(* IEC 61131-3 sources: codesys-api/examples/plc_architecture/st, 45 files *)

(* ---- E_BusFormat.st ---- *)
// How an entry's raw value sits in a block's reply: one bit, or one or two 16-bit registers.
{attribute 'qualified_only'}
{attribute 'strict'}
TYPE E_BusFormat :
(
	SINGLE_BIT := 0,
	INT16 := 1,
	UINT16 := 2,
	INT32 := 3,
	UINT32 := 4,
	FLOAT32 := 5
) USINT;
END_TYPE

(* ---- E_BusFunction.st ---- *)
// Modbus read function of a poll block. Writes (FC06) come from GVL_Bus.Writes.
{attribute 'qualified_only'}
{attribute 'strict'}
TYPE E_BusFunction :
(
	READ_COILS := 1,
	READ_DISCRETE_INPUTS := 2,
	READ_HOLDING_REGISTERS := 3,
	READ_INPUT_REGISTERS := 4
) USINT;
END_TYPE

(* ---- E_CommandResult.st ---- *)
// Outcome of a remote command, sent back to the sender in the acknowledgement. A retry of an id the PLC has
// already answered gets the original result again; it is never applied twice.
{attribute 'qualified_only'}
{attribute 'strict'}
TYPE E_CommandResult :
(
	PENDING := 0,           // parsed, not yet checked
	ACCEPTED := 1,
	MALFORMED := 2,         // not "<id>,<tag>=<number>,<sent_ms>", or a field too long
	UNKNOWN_TAG := 3,
	NOT_WRITABLE := 4,
	OUT_OF_RANGE := 5,      // outside the tag's range, not 0/1 for a BOOL, not whole for an INT, NaN
	TOO_OLD := 6,           // older than allowed, dated in the future, or waited too long in the queue
	OUT_OF_ORDER := 7,      // older than the last command applied to the same tag
	INTERLOCKED := 8,       // a start while not permitted, or sent before the permit came back
	CLOCK_NOT_SYNCED := 9   // the PLC's wall clock isn't plausible, so freshness can't be checked
) USINT;
END_TYPE

(* ---- E_Quality.st ---- *)
// Quality of a tag's value. Interlocks and publishing look at this, not just at the number.
{attribute 'qualified_only'}
{attribute 'strict'}
TYPE E_Quality :
(
	INIT := 0,          // no value since start-up
	GOOD := 1,
	STALE := 2,         // no fresh value from the source within StaleAfter
	COMM_FAIL := 3,     // the source reports a communication error
	INVALID := 4        // out of range, or not computable (e.g. division by zero)
) USINT;
END_TYPE

(* ---- E_TagKind.st ---- *)
{attribute 'qualified_only'}
{attribute 'strict'}
TYPE E_TagKind :
(
	BOOL_TAG := 0,
	INT_TAG := 1,
	REAL_TAG := 2
) USINT;
END_TYPE

(* ---- ST_BusBlock.st ---- *)
// One read request, repeated every PeriodMs: a run of registers or bits of one device. The generator merges a
// device's nearby channels into as few blocks as possible (at most 125 registers or 2,000 bits each).
TYPE ST_BusBlock :
STRUCT
	Line : INT;                         // index in GVL_Bus.Lines
	UnitId : UINT;
	ReadFunction : E_BusFunction;
	Start : UINT;                       // zero-based register or bit address (CODESYS numbering)
	Count : UINT;
	PeriodMs : UDINT := 1000;
	FirstEntry : INT;                   // GVL_Bus.Entries[FirstEntry .. FirstEntry + EntryCount - 1]
	EntryCount : INT;
	Source : INT;                       // the device's source in GVL_Tags (health and age)
END_STRUCT
END_TYPE

(* ---- ST_BusEntry.st ---- *)
// Where one tag's raw value sits in its block's reply. Scaling is the tag's own (ST_TagConfig.Scale and
// Offset); the bus only delivers the device's number.
TYPE ST_BusEntry :
STRUCT
	Offset : UINT;                      // registers (or bits) from the block's Start
	Format : E_BusFormat;
	IsWordSwapped : BOOL;               // 32-bit values: low word first
	HasSentinel : BOOL;                 // a raw value the device uses for "no reading"
	Sentinel : DINT;                    // e.g. -999 for an open thermocouple; delivered as NaN, so the tag is INVALID
	TagIndex : INT;
END_STRUCT
END_TYPE

(* ---- ST_BusLine.st ---- *)
// One Modbus connection: a TCP server (a device or an RS485 gateway port) or one of the PLC's serial ports.
// Every device on it shares this one connection; requests on it run one at a time.
TYPE ST_BusLine :
STRUCT
	IsSerial : BOOL;
	Address : ARRAY[0..3] OF BYTE;      // TCP: server IP
	Port : UINT := 502;                 // TCP: server port
	ComPort : INT := 1;                 // serial: 1 to 4
	RtsControl : USINT;                 // serial: 0 disabled, 1 on, 2 handshake, 3 toggle (RS485 direction)
	Baudrate : UDINT := 9600;           // serial: 9600, 19200, 38400, 57600 or 115200
	Parity : USINT;                     // serial: 0 none, 1 odd, 2 even
	ReplyTimeoutMs : UDINT := 500;
END_STRUCT
END_TYPE

(* ---- ST_BusWrite.st ---- *)
// A writable tag sent to a device register (FC06) when its value changes, and again every RefreshMs so a
// device that restarted gets it back. Raw = (Value - tag Offset) / tag Scale, as a signed 16-bit register.
TYPE ST_BusWrite :
STRUCT
	TagIndex : INT;                     // 0 = unused row
	Line : INT;
	UnitId : UINT;
	Register : UINT;
	RefreshMs : UDINT := 10000;
END_STRUCT
END_TYPE

(* ---- ST_Command.st ---- *)
// One remote command, from the MQTT callback to the control task and back as an acknowledgement.
TYPE ST_Command :
STRUCT
	Id : UDINT;                 // sender's command id, echoed in the acknowledgement
	TagIndex : INT;             // resolved when received; 0 = unknown tag
	Value : REAL;
	SentAtMs : ULINT;           // wall-clock ms from the bridge, the one command sender
	ReceivedAtMs : ULINT;
	Result : E_CommandResult;
END_STRUCT
END_TYPE

(* ---- ST_TagConfig.st ---- *)
// Static description of one tag. Generated from the config sheet into GVL_Tags.TagConfig;
// the program never writes it.
TYPE ST_TagConfig :
STRUCT
	Name : STRING(24);          // tag key, exactly as the bridge layout spells it; sized by the generator from the longest name
	Kind : E_TagKind;
	Scale : REAL := 1.0;        // Value := Raw * Scale + Offset
	Offset : REAL;
	MinValue : REAL;            // a value outside [MinValue, MaxValue], or NaN, is INVALID
	MaxValue : REAL;
	DefaultValue : REAL;        // writable tags start here (alarm setpoints from the sheet; requests 0)
	Deadband : REAL;            // report-by-exception: publish when the value moved more than this
	StaleAfter : TIME := T#5S;  // no fresh value from the source for this long -> STALE
	IsWritable : BOOL;          // may a remote command change it (setpoints, start/stop requests)?
	Source : INT;               // communication source in GVL_Tags.SourceIsHealthy; 0 = local I/O
END_STRUCT
END_TYPE

(* ---- ST_TagState.st ---- *)
// Live state of one tag. Written only by PRG_Control, each field by one step.
TYPE ST_TagState :
STRUCT
	Raw : REAL;                 // step 1: as read from the I/O or the bus
	SourceQuality : E_Quality;  // step 1: from the source's health and age
	Value : REAL;               // step 3 (step 2 for writable tags); BOOL tags use 0.0 / 1.0
	Quality : E_Quality;        // step 3: SourceQuality plus range checks (step 2 for writable tags)
	UpdatedAtMs : ULINT;        // step 1 (step 2 for writable tags): last fresh value, monotonic ms
	LastCommandSentAtMs : ULINT; // step 2: sender time of the last command applied, for ordering
END_STRUCT
END_TYPE

(* ---- GVL_Bus.st ---- *)
// Modbus devices and their hand-over to the control task. Tables are generated from the config sheets'
// rs485Config (and Modbus TCP devices); PRG_Bus (bus task) is the only writer of everything below them.
// Example: AIT-1508 is holding register 40002 (item 1) of RTU unit 24 on the PLC's first serial port.
{attribute 'qualified_only'}
VAR_GLOBAL CONSTANT
	LINE_COUNT : INT := 1;
	BLOCK_COUNT : INT := 1;
	ENTRY_COUNT : INT := 1;
	WRITE_COUNT : INT := 1;
	FAIL_LIMIT : UINT := 3;             // consecutive failed requests before a device is COMM_FAIL
	BACKOFF_MS : UDINT := 5000;         // a failed device is polled this rarely, so it can't slow its line
END_VAR
VAR_GLOBAL
	// Generated; never written by the program.
	Lines : ARRAY[1..LINE_COUNT] OF ST_BusLine := [(IsSerial := TRUE, ComPort := 1, Baudrate := 9600)];
	Blocks : ARRAY[1..BLOCK_COUNT] OF ST_BusBlock := [
		(Line := 1, UnitId := 24, ReadFunction := E_BusFunction.READ_HOLDING_REGISTERS, Start := 1, Count := 1,
		 PeriodMs := 500, FirstEntry := 1, EntryCount := 1, Source := 1)];
	Entries : ARRAY[1..ENTRY_COUNT] OF ST_BusEntry := [(Offset := 0, Format := E_BusFormat.UINT16, TagIndex := 1)];
	Writes : ARRAY[1..WRITE_COUNT] OF ST_BusWrite;          // no device setpoints in this example
	IsBusSource : ARRAY[0..GVL_Tags.SOURCE_COUNT] OF BOOL := [FALSE, TRUE, FALSE];

	// Bus task -> control task. For a source with SourceWriting TRUE the control task was started while the
	// bus task was mid-update: it keeps last scan's values for that source. (Both tasks on one core: control
	// never runs while the bus task writes, except by preempting it.)
	Raw : ARRAY[1..GVL_Tags.TAG_COUNT] OF REAL;             // decoded device numbers, before tag scaling
	SourceWriting : ARRAY[0..GVL_Tags.SOURCE_COUNT] OF BOOL;
	SourceHealthy : ARRAY[0..GVL_Tags.SOURCE_COUNT] OF BOOL := [TRUE, TRUE, TRUE];   // until FAIL_LIMIT failures: INIT, not COMM_FAIL
	SourceLastGoodMs : ARRAY[0..GVL_Tags.SOURCE_COUNT] OF ULINT;   // F_NowMs of the last good reply

	// Diagnostics
	SourceFailCount : ARRAY[0..GVL_Tags.SOURCE_COUNT] OF UINT;
	BlockReads : ARRAY[1..BLOCK_COUNT] OF UDINT;
	BlockErrors : ARRAY[1..BLOCK_COUNT] OF UDINT;
	BlockLastError : ARRAY[1..BLOCK_COUNT] OF UDINT;        // ModbusFB.Error
	BlockLastException : ARRAY[1..BLOCK_COUNT] OF UDINT;    // Modbus exception code
	WriteCount : ARRAY[1..WRITE_COUNT] OF UDINT;
	WriteErrors : ARRAY[1..WRITE_COUNT] OF UDINT;
END_VAR

(* ---- GVL_Tags.st ---- *)
// The tag table and the hand-over points between the control task and the comms task.
// Ownership: every variable below has exactly one writer, named in its comment.
// Changing the table (rows, order, sizes) needs a full download: queued commands and the publisher's
// history refer to rows by index, so an online change must not reinterpret them.
{attribute 'qualified_only'}
VAR_GLOBAL CONSTANT
	TAG_COUNT : INT := 4;               // generated from the config sheet
	SOURCE_COUNT : INT := 2;            // Modbus slaves and remote PLCs; 0 = local I/O
	// Indices for hand-written logic, generated with the table so names and indices stay in step
	TAG_AIT_1508 : INT := 1;
	TAG_AIT_1508_HH_SP : INT := 2;
	TAG_P_1502_REQUEST : INT := 3;
	TAG_LSS_E_STOP : INT := 4;
END_VAR
VAR_GLOBAL
	// Generated from the config sheet; never written by the program.
	TagConfig : ARRAY[1..TAG_COUNT] OF ST_TagConfig := [
		(Name := 'AIT-1508', Kind := E_TagKind.REAL_TAG, Scale := 0.01, MinValue := 0.0, MaxValue := 14.0,
		 Deadband := 0.05, StaleAfter := T#3S, Source := 1),
		(Name := 'AIT-1508_HH_SP', Kind := E_TagKind.REAL_TAG, MinValue := 0.0, MaxValue := 14.0,
		 DefaultValue := 12.5, IsWritable := TRUE),
		(Name := 'P-1502', Kind := E_TagKind.BOOL_TAG, MinValue := 0.0, MaxValue := 1.0, IsWritable := TRUE),
		(Name := 'LSS-E-STOP', Kind := E_TagKind.BOOL_TAG, MinValue := 0.0, MaxValue := 1.0, StaleAfter := T#3S, Source := 2)];

	Tags : ARRAY[1..TAG_COUNT] OF ST_TagState;               // writer: PRG_Control
	RawInputs : ARRAY[1..TAG_COUNT] OF REAL;                  // writer: I/O mapping (control task)
	// Source health and the time of each source's last sample. Writer: the source adapters, which run in the
	// control task (Modbus diagnostics are read there). Data from other tasks (e.g. remote PLCs over MQTT)
	// reaches them through a queue, never by writing these from another task. Not in the skeleton.
	SourceIsHealthy : ARRAY[0..SOURCE_COUNT] OF BOOL := [TRUE, FALSE, FALSE];
	SourceUpdatedAtMs : ARRAY[0..SOURCE_COUNT] OF ULINT;      // 0 = no sample since start-up

	// Control -> comms: a consistent copy of Tags, made when the comms task asks for one.
	PublishSnapshot : ARRAY[1..TAG_COUNT] OF ST_TagState;    // writer: PRG_Control
	SnapshotRequest : UDINT;                                  // writer: PRG_Comms (increments to ask)
	SnapshotSequence : UDINT;                                 // writer: PRG_Control (= SnapshotRequest when served)

	// Comms -> control and back. Each queue has one producer task and one consumer task.
	// Both tasks must run on the same core, or the queues need the target's atomics and barriers.
	Commands : FB_CommandQueue;         // Push: FB_CommandReceiver (comms task); Pop: PRG_Control
	Acks : FB_CommandQueue;             // Push: PRG_Control; Pop: PRG_Comms

	// Physical outputs, mapped to I/O.
	P_1502_RUN : BOOL;                  // writer: PRG_Control.WriteOutputs, nothing else
END_VAR

(* ---- F_BusDecode.st ---- *)
FUNCTION F_BusDecode : BOOL
// Turns one block's reply into GVL_Bus.Raw for each of its entries. Call it with the source's SourceWriting
// flag set. A sentinel ("no reading") becomes NaN, so the tag goes INVALID in ComputeValues. Independent of
// the transport: FB_BusLine passes a ModbusFB reply, a native device-tree channel its mapped input image.
VAR_INPUT
	FirstEntry : INT;
	EntryCount : INT;
END_VAR
VAR_IN_OUT
	Words : ARRAY[0..124] OF WORD;      // register reply, first register at index 0
	Bits : ARRAY[0..1999] OF BYTE;      // bit reply, one byte per bit
END_VAR
VAR
	Index : INT;
	Entry : ST_BusEntry;
	RawInt : DINT;
	Raw32 : DWORD;
	Value : REAL;
	pReal : POINTER TO REAL;
	NanBits : DWORD := 16#7FC00000;
END_VAR
// ---- implementation ----
FOR Index := FirstEntry TO FirstEntry + EntryCount - 1 DO
	Entry := GVL_Bus.Entries[Index];
	IF Entry.Format = E_BusFormat.SINGLE_BIT THEN
		RawInt := SEL(Bits[Entry.Offset] <> 0, 0, 1);   // ModbusFB unpacks bit replies: one byte per coil (bench, 2026-10-20)
		Value := DINT_TO_REAL(RawInt);
	ELSIF Entry.Format = E_BusFormat.INT16 THEN
		RawInt := INT_TO_DINT(WORD_TO_INT(Words[Entry.Offset]));
		Value := DINT_TO_REAL(RawInt);
	ELSIF Entry.Format = E_BusFormat.UINT16 THEN
		RawInt := WORD_TO_DINT(Words[Entry.Offset]);
		Value := DINT_TO_REAL(RawInt);
	ELSE
		IF Entry.IsWordSwapped THEN
			Raw32 := SHL(WORD_TO_DWORD(Words[Entry.Offset + 1]), 16) OR WORD_TO_DWORD(Words[Entry.Offset]);
		ELSE
			Raw32 := SHL(WORD_TO_DWORD(Words[Entry.Offset]), 16) OR WORD_TO_DWORD(Words[Entry.Offset + 1]);
		END_IF
		RawInt := DWORD_TO_DINT(Raw32);
		IF Entry.Format = E_BusFormat.FLOAT32 THEN
			pReal := ADR(Raw32);
			Value := pReal^;
		ELSIF Entry.Format = E_BusFormat.UINT32 THEN
			Value := UDINT_TO_REAL(DWORD_TO_UDINT(Raw32));
		ELSE
			Value := DINT_TO_REAL(RawInt);
		END_IF
	END_IF
	IF Entry.HasSentinel AND RawInt = Entry.Sentinel THEN
		pReal := ADR(NanBits);
		Value := pReal^;
	END_IF
	GVL_Bus.Raw[Entry.TagIndex] := Value;
END_FOR
F_BusDecode := TRUE;

(* ---- F_FindTag.st ---- *)
FUNCTION F_FindTag : INT
// Index of the tag with this name, 0 if there is none. A linear search is fine for occasional commands;
// with thousands of tags and frequent commands, generate the table sorted by name and search it binarily.
VAR_INPUT
	Name : STRING(24);
END_VAR
VAR
	Index : INT;
END_VAR
// ---- implementation ----
F_FindTag := 0;
FOR Index := 1 TO GVL_Tags.TAG_COUNT DO
	IF GVL_Tags.TagConfig[Index].Name = Name THEN
		F_FindTag := Index;
		RETURN;
	END_IF
END_FOR

(* ---- F_IsNumberText.st ---- *)
FUNCTION F_IsNumberText : BOOL
// TRUE for a plain decimal number of 1..MaxLength characters: an optional leading '-', digits, at most one
// '.'. With IsDigitsOnly, only unsigned integers (ids, timestamps). MaxLength keeps the value inside the
// target type (9 digits for a UDINT id, 15 for a millisecond timestamp). Run this before STRING_TO_REAL/
// _UDINT/_ULINT, which return 0 for text they can't read.
VAR_INPUT
	Text : STRING(40);
	IsDigitsOnly : BOOL;
	MaxLength : INT;
END_VAR
VAR
	pChar : POINTER TO BYTE;
	Length : INT;
	Index : INT;
	Digits : INT;
	Dots : INT;
END_VAR
// ---- implementation ----
F_IsNumberText := FALSE;
Length := LEN(Text);
IF Length < 1 OR Length > MaxLength THEN
	RETURN;
END_IF
pChar := ADR(Text);
FOR Index := 0 TO Length - 1 DO
	IF pChar[Index] >= 16#30 AND pChar[Index] <= 16#39 THEN
		Digits := Digits + 1;
	ELSIF pChar[Index] = 16#2E AND NOT IsDigitsOnly THEN
		Dots := Dots + 1;
	ELSIF NOT (pChar[Index] = 16#2D AND Index = 0 AND NOT IsDigitsOnly) THEN
		RETURN;                         // any other character, or '-' anywhere but first
	END_IF
END_FOR
F_IsNumberText := Digits > 0 AND Dots <= 1;

(* ---- F_NowMs.st ---- *)
FUNCTION F_NowMs : ULINT
// Monotonic milliseconds since start-up, for ages and timeouts. Not wall-clock time.
VAR
	Microseconds : ULINT;
END_VAR
// ---- implementation ----
SysTimeCore.SysTimeGetUs(pUsTime := Microseconds);
F_NowMs := Microseconds / 1000;

(* ---- F_NowUs.st ---- *)
FUNCTION F_NowUs : ULINT
// Monotonic microseconds since start-up, for time budgets within a scan. Not wall-clock time.
VAR
	Microseconds : ULINT;
END_VAR
// ---- implementation ----
SysTimeCore.SysTimeGetUs(pUsTime := Microseconds);
F_NowUs := Microseconds;

(* ---- F_WallClockMs.st ---- *)
FUNCTION F_WallClockMs : ULINT
// Milliseconds since 1970 from the controller's real-time clock, to compare with senders' timestamps.
// Only meaningful while the clock is synchronized (SNTP).
VAR
	Timestamp : ULINT;
END_VAR
// ---- implementation ----
SysTimeRtc.SysTimeRtcHighResGet(pTimestamp := Timestamp);
F_WallClockMs := Timestamp;

(* ---- FB_BusLine.st ---- *)
{attribute 'no_assign'}
FUNCTION_BLOCK FB_BusLine
// One Modbus connection (GVL_Bus.Lines[LineIndex]) with every block and write on it. Called every bus-task
// cycle. One request is in flight at a time; the next starts in the same call that finishes the last
// (ModbusFB's "daisy chain"), so the line never idles a task cycle between requests.
VAR_INPUT
	LineIndex : INT;
	IsEnabled : BOOL := TRUE;
	Reconnect : BOOL;                   // rising edge: drop the connection and connect with the current settings
END_VAR
VAR_OUTPUT
	IsConnected : BOOL;
	RequestCount : UDINT;
	ErrorCount : UDINT;
	LastRequestUs : UDINT;              // start to reply of the last request
	MaxRequestUs : UDINT;
END_VAR
VAR
	ClientTcp : ModbusFB.ClientTCP;
	ClientRtu : ModbusFB.ClientSerial;
	Client : REFERENCE TO ModbusFB.Client;   // whichever of the two this line uses (set by CallClient)
	ReadCoils : ModbusFB.ClientRequestReadCoils;
	ReadDiscrete : ModbusFB.ClientRequestReadDiscreteInputs;
	ReadHolding : ModbusFB.ClientRequestReadHoldingRegisters;
	ReadInput : ModbusFB.ClientRequestReadInputRegisters;
	WriteRegister : ModbusFB.ClientRequestWriteSingleRegister;
	Words : ARRAY[0..124] OF WORD;      // reply of the active register block
	Bits : ARRAY[0..1999] OF BYTE;      // reply of the active bit block: one byte per bit (ModbusFB unpacks them)
	Block : ST_BusBlock;                // copy of the active block
	ActiveBlock : INT;                  // 0 = no read in flight
	ActiveWrite : INT;                  // 0 = no write in flight
	NextBlock : INT := 1;               // round-robin start
	BlockDueMs : ARRAY[1..GVL_Bus.BLOCK_COUNT] OF ULINT;
	WriteDueMs : ARRAY[1..GVL_Bus.WRITE_COUNT] OF ULINT;
	WriteSentValue : ARRAY[1..GVL_Bus.WRITE_COUNT] OF REAL;
	HasWritten : ARRAY[1..GVL_Bus.WRITE_COUNT] OF BOOL;
	WriteValue : REAL;
	WriteRaw : INT;
	IsDone : BOOL;
	IsError : BOOL;
	ErrorId : UDINT;
	Exception : UDINT;
	NowMs : ULINT;
	StartUs : ULINT;
	ReconnectEdge : R_TRIG;
	HoldUntilMs : ULINT;                // connection held down until then (reconnect, client error)
END_VAR
// ---- implementation ----
NowMs := F_NowMs();
ReconnectEdge(CLK := Reconnect);
IF ReconnectEdge.Q THEN
	HoldUntilMs := NowMs + 500;
END_IF
CallClient();

IF ActiveBlock <> 0 OR ActiveWrite <> 0 THEN
	IF CallRequest(IsExecute := TRUE) THEN
		FinishRequest();
	END_IF
END_IF
IF ActiveBlock = 0 AND ActiveWrite = 0 AND IsConnected THEN
	StartNext();
END_IF

(* ---- FB_CommandQueue.st ---- *)
FUNCTION_BLOCK FB_CommandQueue
// Single-producer / single-consumer ring buffer between two tasks. Push is called from one task
// only, Pop from one other task only; each side writes only its own index, so no lock is needed. Push fills
// the slot before it advances Head, so Pop never sees a half-written item. This relies on both tasks running
// on one core; across cores, the index updates need the runtime's atomic operations and memory barriers.
// Usable capacity is SIZE - 1 (one slot stays empty to tell "full" from "empty").
VAR CONSTANT
	SIZE : UINT := 32;
END_VAR
VAR_OUTPUT
	OverflowCount : UDINT;              // items dropped because the queue was full
END_VAR
VAR
	Items : ARRAY[0..SIZE - 1] OF ST_Command;
	Head : UINT;                        // next free slot; written only by Push
	Tail : UINT;                        // next item to take; written only by Pop
END_VAR
// ---- implementation ----
// Everything happens in the Push and Pop methods.

(* ---- FB_CommandReceiver.st ---- *)
FUNCTION_BLOCK FB_CommandReceiver IMPLEMENTS MQTT.MQTT_SUBSCRIBE_CALLBACK
// MQTT subscription callback: turns every received command into an ST_Command and queues it for the
// control task, instead of keeping only the latest message. Runs in the comms task (inside the MQTT client).
// Message format: <id>,<tag>=<value>,<sent_ms>   e.g. '1042,P-1502=1,1769612037947'
VAR_OUTPUT
	ReceivedCount : UDINT;
	MalformedCount : UDINT;
	DroppedCount : UDINT;               // queue full: no acknowledgement, so the sender retries
END_VAR
VAR
	Line : STRING(255);
END_VAR
// ---- implementation ----
// Everything happens in PublishReceived, called by the MQTT library for each message.

(* ---- FB_BusLine.CallClient.st ---- *)
METHOD CallClient : BOOL
// Runs this line's client (TCP or serial) and returns IsConnected. Settings are read when it connects. A client
// error holds the connection down for a second before the next attempt.
VAR
	Port : SysCom.SYS_COM_PORTS;
	Baudrate : SysCom.SYS_COM_BAUDRATE;
	Parity : SysCom.SYS_COM_PARITY;
	Rts : SysCom.SYS_COM_RTS_CONTROL;
END_VAR
// ---- implementation ----
IF GVL_Bus.Lines[LineIndex].IsSerial THEN
	CASE GVL_Bus.Lines[LineIndex].ComPort OF
		2: Port := SysCom.SYS_COM_PORTS.SYS_COMPORT2;
		3: Port := SysCom.SYS_COM_PORTS.SYS_COMPORT3;
		4: Port := SysCom.SYS_COM_PORTS.SYS_COMPORT4;
	ELSE
		Port := SysCom.SYS_COM_PORTS.SYS_COMPORT1;
	END_CASE
	CASE GVL_Bus.Lines[LineIndex].RtsControl OF
		1: Rts := SysCom.SYS_COM_RTS_CONTROL.SYS_RTS_CONTROL_ENABLE;
		2: Rts := SysCom.SYS_COM_RTS_CONTROL.SYS_RTS_CONTROL_HANDSHAKE;
		3: Rts := SysCom.SYS_COM_RTS_CONTROL.SYS_RTS_CONTROL_TOGGLE;
	ELSE
		Rts := SysCom.SYS_COM_RTS_CONTROL.SYS_RTS_CONTROL_DISABLE;
	END_CASE
	CASE GVL_Bus.Lines[LineIndex].Baudrate OF
		19200: Baudrate := SysCom.SYS_COM_BAUDRATE.SYS_BR_19200;
		38400: Baudrate := SysCom.SYS_COM_BAUDRATE.SYS_BR_38400;
		57600: Baudrate := SysCom.SYS_COM_BAUDRATE.SYS_BR_57600;
		115200: Baudrate := SysCom.SYS_COM_BAUDRATE.SYS_BR_115200;
	ELSE
		Baudrate := SysCom.SYS_COM_BAUDRATE.SYS_BR_9600;
	END_CASE
	CASE GVL_Bus.Lines[LineIndex].Parity OF
		1: Parity := SysCom.SYS_COM_PARITY.SYS_ODDPARITY;
		2: Parity := SysCom.SYS_COM_PARITY.SYS_EVENPARITY;
	ELSE
		Parity := SysCom.SYS_COM_PARITY.SYS_NOPARITY;
	END_CASE
	Client REF= ClientRtu;
	ClientRtu(xConnect := IsEnabled AND NowMs >= HoldUntilMs, iPort := Port, dwBaudrate := Baudrate, eParity := Parity,
		eRTScontrol := Rts);
	IsConnected := ClientRtu.xConnected;
	IF ClientRtu.xError AND NowMs >= HoldUntilMs THEN
		HoldUntilMs := NowMs + 1000;
	END_IF
ELSE
	Client REF= ClientTcp;
	ClientTcp(xConnect := IsEnabled AND NowMs >= HoldUntilMs, aIPaddr := GVL_Bus.Lines[LineIndex].Address,
		uiPort := GVL_Bus.Lines[LineIndex].Port, tConnnectTimeOut := T#2S);
	IsConnected := ClientTcp.xConnected;
	IF ClientTcp.xError AND NowMs >= HoldUntilMs THEN
		HoldUntilMs := NowMs + 1000;
	END_IF
END_IF
CallClient := IsConnected;

(* ---- FB_BusLine.CallRequest.st ---- *)
METHOD CallRequest : BOOL
// Calls the request block of the active read or write. TRUE when it finished (IsDone or IsError). Called with
// IsExecute FALSE once afterwards: the falling edge that lets the same request block start again.
VAR_INPUT
	IsExecute : BOOL;
END_VAR
VAR
	ReplyUs : UDINT;
	TimeoutUs : UDINT;
END_VAR
// ---- implementation ----
ReplyUs := GVL_Bus.Lines[LineIndex].ReplyTimeoutMs * 1000;
TimeoutUs := ReplyUs + 1000000;
IF ActiveWrite <> 0 THEN
	WriteRegister(rClient := Client, xExecute := IsExecute, uiUnitId := GVL_Bus.Writes[ActiveWrite].UnitId,
		uiItem := GVL_Bus.Writes[ActiveWrite].Register, uiValue := INT_TO_UINT(WriteRaw),
		udiReplyTimeout := ReplyUs, udiTimeOut := TimeoutUs, uiMaxRetries := 0);
	IsDone := WriteRegister.xDone;
	IsError := WriteRegister.xError;
	ErrorId := TO_UDINT(WriteRegister.eErrorID);
	Exception := TO_UDINT(WriteRegister.eException);
ELSIF Block.ReadFunction = E_BusFunction.READ_HOLDING_REGISTERS THEN
	ReadHolding(rClient := Client, xExecute := IsExecute, uiUnitId := Block.UnitId, uiStartItem := Block.Start,
		uiQuantity := Block.Count, pData := ADR(Words), udiReplyTimeout := ReplyUs, udiTimeOut := TimeoutUs, uiMaxRetries := 0);
	IsDone := ReadHolding.xDone;
	IsError := ReadHolding.xError;
	ErrorId := TO_UDINT(ReadHolding.eErrorID);
	Exception := TO_UDINT(ReadHolding.eException);
ELSIF Block.ReadFunction = E_BusFunction.READ_INPUT_REGISTERS THEN
	ReadInput(rClient := Client, xExecute := IsExecute, uiUnitId := Block.UnitId, uiStartItem := Block.Start,
		uiQuantity := Block.Count, pData := ADR(Words), udiReplyTimeout := ReplyUs, udiTimeOut := TimeoutUs, uiMaxRetries := 0);
	IsDone := ReadInput.xDone;
	IsError := ReadInput.xError;
	ErrorId := TO_UDINT(ReadInput.eErrorID);
	Exception := TO_UDINT(ReadInput.eException);
ELSIF Block.ReadFunction = E_BusFunction.READ_COILS THEN
	ReadCoils(rClient := Client, xExecute := IsExecute, uiUnitId := Block.UnitId, uiStartItem := Block.Start,
		uiQuantity := Block.Count, pData := ADR(Bits), udiReplyTimeout := ReplyUs, udiTimeOut := TimeoutUs, uiMaxRetries := 0);
	IsDone := ReadCoils.xDone;
	IsError := ReadCoils.xError;
	ErrorId := TO_UDINT(ReadCoils.eErrorID);
	Exception := TO_UDINT(ReadCoils.eException);
ELSE
	ReadDiscrete(rClient := Client, xExecute := IsExecute, uiUnitId := Block.UnitId, uiStartItem := Block.Start,
		uiQuantity := Block.Count, pData := ADR(Bits), udiReplyTimeout := ReplyUs, udiTimeOut := TimeoutUs, uiMaxRetries := 0);
	IsDone := ReadDiscrete.xDone;
	IsError := ReadDiscrete.xError;
	ErrorId := TO_UDINT(ReadDiscrete.eErrorID);
	Exception := TO_UDINT(ReadDiscrete.eException);
END_IF
CallRequest := IsDone OR IsError;

(* ---- FB_BusLine.FinishRequest.st ---- *)
METHOD FinishRequest : BOOL
// The active request finished: take its result, update the device's health and schedule the block again.
// A device that failed FAIL_LIMIT times in a row is COMM_FAIL and polled only every BACKOFF_MS.
VAR
	Source : INT;
END_VAR
// ---- implementation ----
LastRequestUs := ULINT_TO_UDINT(F_NowUs() - StartUs);
MaxRequestUs := MAX(MaxRequestUs, LastRequestUs);
RequestCount := RequestCount + 1;
IF IsError THEN
	ErrorCount := ErrorCount + 1;
END_IF

IF ActiveWrite <> 0 THEN
	IF IsDone THEN
		GVL_Bus.WriteCount[ActiveWrite] := GVL_Bus.WriteCount[ActiveWrite] + 1;
		WriteDueMs[ActiveWrite] := NowMs + GVL_Bus.Writes[ActiveWrite].RefreshMs;
	ELSE
		GVL_Bus.WriteErrors[ActiveWrite] := GVL_Bus.WriteErrors[ActiveWrite] + 1;
		WriteDueMs[ActiveWrite] := NowMs + 1000;     // retried in a second, not every call
	END_IF
	HasWritten[ActiveWrite] := TRUE;
	WriteSentValue[ActiveWrite] := WriteValue;
	CallRequest(IsExecute := FALSE);
	ActiveWrite := 0;
	FinishRequest := TRUE;
	RETURN;
END_IF

Source := Block.Source;
IF IsDone THEN
	GVL_Bus.SourceWriting[Source] := TRUE;
	F_BusDecode(FirstEntry := Block.FirstEntry, EntryCount := Block.EntryCount, Words := Words, Bits := Bits);
	GVL_Bus.SourceLastGoodMs[Source] := NowMs;
	GVL_Bus.SourceHealthy[Source] := TRUE;
	GVL_Bus.SourceFailCount[Source] := 0;
	GVL_Bus.SourceWriting[Source] := FALSE;
	GVL_Bus.BlockReads[ActiveBlock] := GVL_Bus.BlockReads[ActiveBlock] + 1;
	BlockDueMs[ActiveBlock] := NowMs + Block.PeriodMs;
ELSE
	GVL_Bus.BlockErrors[ActiveBlock] := GVL_Bus.BlockErrors[ActiveBlock] + 1;
	GVL_Bus.BlockLastError[ActiveBlock] := ErrorId;
	GVL_Bus.BlockLastException[ActiveBlock] := Exception;
	IF GVL_Bus.SourceFailCount[Source] < 65535 THEN
		GVL_Bus.SourceFailCount[Source] := GVL_Bus.SourceFailCount[Source] + 1;
	END_IF
	IF GVL_Bus.SourceFailCount[Source] >= GVL_Bus.FAIL_LIMIT THEN
		GVL_Bus.SourceWriting[Source] := TRUE;
		GVL_Bus.SourceHealthy[Source] := FALSE;
		GVL_Bus.SourceWriting[Source] := FALSE;
		BlockDueMs[ActiveBlock] := NowMs + MAX(Block.PeriodMs, GVL_Bus.BACKOFF_MS);
	ELSE
		BlockDueMs[ActiveBlock] := NowMs + Block.PeriodMs;
	END_IF
END_IF
CallRequest(IsExecute := FALSE);
ActiveBlock := 0;
FinishRequest := TRUE;

(* ---- FB_BusLine.StartNext.st ---- *)
METHOD StartNext : BOOL
// Starts the next request on this line, TRUE if it started one. Writes go first, so a changed setpoint never
// waits behind a round of reads. Reads go round-robin over the due blocks, so one device can't starve another.
VAR
	Index : INT;
	Candidate : INT;
	TagIndex : INT;
	RawValue : REAL;
END_VAR
// ---- implementation ----
FOR Index := 1 TO GVL_Bus.WRITE_COUNT DO
	TagIndex := GVL_Bus.Writes[Index].TagIndex;
	IF TagIndex > 0 AND GVL_Bus.Writes[Index].Line = LineIndex
			AND_THEN GVL_Tags.Tags[TagIndex].Quality = E_Quality.GOOD
			AND_THEN (NOT HasWritten[Index] OR GVL_Tags.Tags[TagIndex].Value <> WriteSentValue[Index] OR NowMs >= WriteDueMs[Index]) THEN
		WriteValue := GVL_Tags.Tags[TagIndex].Value;
		RawValue := (WriteValue - GVL_Tags.TagConfig[TagIndex].Offset) / GVL_Tags.TagConfig[TagIndex].Scale;
		// Range first, conversion after: REAL_TO_INT outside INT can fault.
		IF RawValue >= -32768.0 AND RawValue <= 32767.0 THEN
			WriteRaw := REAL_TO_INT(RawValue);
			ActiveWrite := Index;
			StartUs := F_NowUs();
			CallRequest(IsExecute := TRUE);
			StartNext := TRUE;
			RETURN;
		END_IF
		GVL_Bus.WriteErrors[Index] := GVL_Bus.WriteErrors[Index] + 1;
		HasWritten[Index] := TRUE;              // don't retry an unwritable value every call
		WriteSentValue[Index] := WriteValue;
		WriteDueMs[Index] := NowMs + GVL_Bus.Writes[Index].RefreshMs;
	END_IF
END_FOR

FOR Index := 0 TO GVL_Bus.BLOCK_COUNT - 1 DO
	Candidate := (NextBlock - 1 + Index) MOD GVL_Bus.BLOCK_COUNT + 1;
	IF GVL_Bus.Blocks[Candidate].Line = LineIndex AND NowMs >= BlockDueMs[Candidate] THEN
		ActiveBlock := Candidate;
		Block := GVL_Bus.Blocks[Candidate];
		NextBlock := Candidate MOD GVL_Bus.BLOCK_COUNT + 1;
		StartUs := F_NowUs();
		CallRequest(IsExecute := TRUE);
		StartNext := TRUE;
		RETURN;
	END_IF
END_FOR

(* ---- FB_CommandQueue.Pop.st ---- *)
METHOD Pop : BOOL
VAR_IN_OUT
	Item : ST_Command;
END_VAR
// ---- implementation ----
IF Tail = Head THEN
	Pop := FALSE;
	RETURN;
END_IF
Item := Items[Tail];
Tail := (Tail + 1) MOD SIZE;
Pop := TRUE;

(* ---- FB_CommandQueue.Push.st ---- *)
METHOD Push : BOOL
VAR_INPUT
	Item : ST_Command;
END_VAR
VAR
	Next : UINT;
END_VAR
// ---- implementation ----
Next := (Head + 1) MOD SIZE;
IF Next = Tail THEN
	OverflowCount := OverflowCount + 1;
	Push := FALSE;
	RETURN;
END_IF
Items[Head] := Item;
Head := Next;                           // publish the item only once it is complete
Push := TRUE;

(* ---- FB_CommandReceiver.PublishReceived.st ---- *)
METHOD PublishReceived : BOOL
VAR_INPUT
	Data : MQTT.CALLBACK_DATA;
END_VAR
VAR
	Command : ST_Command;
	Rest : STRING(255);
	IdText : STRING(40);
	ValueText : STRING(40);
	TimeText : STRING(40);
	FirstComma : INT;
	EqualsAt : INT;
	SecondComma : INT;
END_VAR
// ---- implementation ----
// Copy the payload now: the library reuses its buffer for the next message. The copy stops at SIZEOF(Line);
// the length test below rejects a message that was cut short or holds a NUL.
Line := Data.PayloadString^;
ReceivedCount := ReceivedCount + 1;
Command.ReceivedAtMs := F_NowMs();
Command.Result := E_CommandResult.MALFORMED;

// Keep the id whenever it is readable, so even a malformed command gets an answer the sender can match.
FirstComma := FIND(Line, ',');
IF FirstComma > 1 THEN
	IdText := LEFT(Line, FirstComma - 1);
	IF F_IsNumberText(Text := IdText, IsDigitsOnly := TRUE, MaxLength := 9) THEN
		Command.Id := STRING_TO_UDINT(IdText);
	END_IF
END_IF

EqualsAt := FIND(Line, '=');
Rest := RIGHT(Line, LEN(Line) - EqualsAt);
SecondComma := FIND(Rest, ',');
ValueText := LEFT(Rest, SecondComma - 1);
TimeText := RIGHT(Rest, LEN(Rest) - SecondComma);
IF Data.PayloadSize = INT_TO_UDINT(LEN(Line)) AND Command.Id <> 0 AND EqualsAt > FirstComma + 1 AND SecondComma > 1
		AND F_IsNumberText(Text := ValueText, IsDigitsOnly := FALSE, MaxLength := 15)
		AND F_IsNumberText(Text := TimeText, IsDigitsOnly := TRUE, MaxLength := 15) THEN
	Command.TagIndex := F_FindTag(Name := MID(Line, EqualsAt - FirstComma - 1, FirstComma + 1));
	Command.Value := STRING_TO_REAL(ValueText);
	Command.SentAtMs := STRING_TO_ULINT(TimeText);
	Command.Result := E_CommandResult.PENDING;
ELSE
	MalformedCount := MalformedCount + 1;   // still queued: the control task (the only Acks producer) answers it
END_IF

IF NOT GVL_Tags.Commands.Push(Item := Command) THEN
	DroppedCount := DroppedCount + 1;       // no answer: the sender times out and retries with the same id
END_IF
PublishReceived := TRUE;

(* ---- PRG_Bus.st ---- *)
PROGRAM PRG_Bus
// Bus task: fast cycle (about 5 ms), priority between PRG_Control and PRG_Comms. Owns every Modbus connection;
// the control task only sees GVL_Bus.Raw and the per-source health, through CollectBusInputs.
VAR
	Lines : ARRAY[1..GVL_Bus.LINE_COUNT] OF FB_BusLine;
	Reconnect : ARRAY[1..GVL_Bus.LINE_COUNT] OF BOOL;   // set online to reconnect a line with new settings
	Index : INT;
END_VAR
// ---- implementation ----
FOR Index := 1 TO GVL_Bus.LINE_COUNT DO
	Lines[Index](LineIndex := Index, Reconnect := Reconnect[Index]);
	Reconnect[Index] := FALSE;
END_FOR

(* ---- PRG_Comms.AppendTag.st ---- *)
// Action AppendTag: tag number Index as a "name:value" line, if it changed beyond its deadband, its quality
// changed, or this is a full refresh. The history is not touched here: CommitSent moves it on once the
// message is out. Until quality has its own field on the wire (an open decision, see the design), a tag
// that isn't GOOD is sent as NaN, never as a converted number.
// ---- implementation ----
TagValue := GVL_Tags.PublishSnapshot[Index].Value;
IF IsFullRefresh
		OR GVL_Tags.PublishSnapshot[Index].Quality <> LastSentQuality[Index]
		OR ABS(TagValue - LastSentValue[Index]) > GVL_Tags.TagConfig[Index].Deadband THEN
	// The range test is FALSE for NaN and infinity, and keeps the conversions below inside DINT.
	IF GVL_Tags.PublishSnapshot[Index].Quality <> E_Quality.GOOD OR NOT (TagValue >= -1.0E9 AND TagValue <= 1.0E9) THEN
		ValueText := 'NaN';
	ELSIF GVL_Tags.TagConfig[Index].Kind = E_TagKind.BOOL_TAG THEN
		ValueText := SEL(TagValue > 0.5, '0', '1');
	ELSIF GVL_Tags.TagConfig[Index].Kind = E_TagKind.INT_TAG THEN
		ValueText := DINT_TO_STRING(REAL_TO_DINT(TagValue));
	ELSIF ABS(TagValue) < 1.0E6 THEN    // two decimals: shorter text, and TRUNC stays inside DINT
		ValueText := REAL_TO_STRING(DINT_TO_REAL(TRUNC(TagValue * 100.0 + SEL(TagValue >= 0.0, -0.5, 0.5))) / 100.0);
	ELSE
		ValueText := REAL_TO_STRING(TagValue);
	END_IF
	IsBuildOk := IsBuildOk
		AND_THEN AppendZ(pBuffer := ADR(Payload), Capacity := SIZEOF(Payload), pText := ADR(GVL_Tags.TagConfig[Index].Name), Used := Used)
		AND_THEN AppendZ(pBuffer := ADR(Payload), Capacity := SIZEOF(Payload), pText := ADR(':'), Used := Used)
		AND_THEN AppendZ(pBuffer := ADR(Payload), Capacity := SIZEOF(Payload), pText := ADR(ValueText), Used := Used)
		AND_THEN AppendZ(pBuffer := ADR(Payload), Capacity := SIZEOF(Payload), pText := ADR('$N'), Used := Used);
	IsInMessage[Index] := TRUE;
END_IF

(* ---- PRG_Comms.CommitSent.st ---- *)
// Action CommitSent: the message went out, so its tags' values become the report-by-exception history.
// The snapshot is unchanged until the next request, so it still holds exactly what was sent.
// ---- implementation ----
FOR Index := 1 TO GVL_Tags.TAG_COUNT DO
	IF IsInMessage[Index] THEN
		LastSentValue[Index] := GVL_Tags.PublishSnapshot[Index].Value;
		LastSentQuality[Index] := GVL_Tags.PublishSnapshot[Index].Quality;
		IsInMessage[Index] := FALSE;
	END_IF
END_FOR

(* ---- PRG_Comms.ForgetMessage.st ---- *)
// Action ForgetMessage: the message was too big to build, so nothing was sent. Keep the history as it was
// and make the next message a full refresh, so nothing that changed is lost.
// ---- implementation ----
FOR Index := 1 TO GVL_Tags.TAG_COUNT DO
	IsInMessage[Index] := FALSE;
END_FOR
IsForceFullRefresh := TRUE;

(* ---- PRG_Comms.PublishAcks.st ---- *)
// Action PublishAcks: answer commands as "<id>:<result>" lines, several per message. A batch stays until
// the broker confirms it (QoS 1); the library resends it after a reconnect, so an answer is never dropped here.
// ---- implementation ----
IF NOT IsAckBatchReady AND MqttLink.BROKER_CONNECTED THEN
	AckUsed := 0;
	AckPayload := '';
	WHILE AckUsed < 900 AND_THEN GVL_Tags.Acks.Pop(Item := Ack) DO
		AckLine := CONCAT(CONCAT(UDINT_TO_STRING(Ack.Id), ':'), USINT_TO_STRING(TO_USINT(Ack.Result)));
		AppendZ(pBuffer := ADR(AckPayload), Capacity := SIZEOF(AckPayload), pText := ADR(AckLine), Used := AckUsed);
		AppendZ(pBuffer := ADR(AckPayload), Capacity := SIZEOF(AckPayload), pText := ADR('$N'), Used := AckUsed);
	END_WHILE
	IsAckBatchReady := AckUsed > 0;
END_IF

// Same publisher rules as PublishData: re-arm between sends, keep the batch until done.
IF IsAckBatchReady AND NOT IsAckRequested AND IsAckPublisherArmed THEN
	IsAckRequested := TRUE;
END_IF
AckPublisher(Topic := ADR(TopicAcks), PayloadString := ADR(AckPayload), PublishAsString := TRUE,
	QoSIn := MQTT.QoS.AtLeastOnce, MRetain := FALSE, send := IsAckRequested);
IsAckPublisherArmed := NOT IsAckRequested;
IF AckPublisher.done THEN
	IsAckRequested := FALSE;
	IsAckBatchReady := FALSE;           // confirmed: the next batch can be built
END_IF

(* ---- PRG_Comms.PublishData.st ---- *)
// Action PublishData: once a second, ask the control task for a snapshot, build the message from it over
// several calls (changed tags only, plus a full refresh now and then), and publish it as one message.
// ---- implementation ----
ConnectedEdge(CLK := MqttLink.BROKER_CONNECTED);
IF ConnectedEdge.Q THEN
	IsForceFullRefresh := TRUE;         // the bridge may have missed messages while we were away
END_IF

PublishTimer(IN := NOT PublishTimer.Q, PT := T#1S);
IF PublishTimer.Q AND MqttLink.BROKER_CONNECTED
		AND NOT (IsWaitingForSnapshot OR IsBuilding OR IsMessageReady OR IsRequested) THEN
	GVL_Tags.SnapshotRequest := GVL_Tags.SnapshotRequest + 1;
	IsWaitingForSnapshot := TRUE;
END_IF

IF IsWaitingForSnapshot AND GVL_Tags.SnapshotSequence = GVL_Tags.SnapshotRequest THEN
	IsWaitingForSnapshot := FALSE;
	PublishCount := PublishCount + 1;
	IsFullRefresh := IsForceFullRefresh OR (PublishCount MOD FULL_REFRESH_EVERY) = 1;
	IsForceFullRefresh := FALSE;        // set again by a reconnect or a message that didn't fit
	Used := 0;
	Payload := '';
	IsBuildOk := TRUE;
	NextTag := 1;
	IsBuilding := TRUE;
END_IF

IF IsBuilding THEN
	LastTag := MIN(GVL_Tags.TAG_COUNT, NextTag + TAGS_PER_CALL - 1);
	FOR Index := NextTag TO LastTag DO
		AppendTag();
	END_FOR
	NextTag := LastTag + 1;
	IF NextTag > GVL_Tags.TAG_COUNT THEN
		IsBuilding := FALSE;
		IF NOT IsBuildOk THEN
			ForgetMessage();            // didn't fit: send nothing, try a full message next time
		ELSE
			IsMessageReady := Used > 0; // nothing changed: nothing to send
		END_IF
	END_IF
END_IF

// MQTTPublish starts on a rising edge of send, so it must see FALSE between two messages. Once started, the
// library keeps the request until the broker has it (it resends after a reconnect) and reads Payload through
// its pointer the whole time, so Payload, the snapshot and IsInMessage stay untouched until done.
// SendTimeout only says it is taking long: it does not end the request.
IF IsMessageReady AND NOT IsRequested AND IsPublisherArmed THEN
	IsRequested := TRUE;
END_IF
Publisher(Topic := ADR(TopicData), PayloadString := ADR(Payload), PublishAsString := TRUE,
	QoSIn := MQTT.QoS.AtMostOnce, MRetain := FALSE, send := IsRequested);
IsPublisherArmed := NOT IsRequested;
IF Publisher.done THEN
	IsRequested := FALSE;
	IsMessageReady := FALSE;
	CommitSent();                       // only now does the history move on
END_IF
SlowPublishEdge(CLK := Publisher.SendTimeout);
IF SlowPublishEdge.Q THEN
	SlowPublishCount := SlowPublishCount + 1;
END_IF

(* ---- PRG_Comms.st ---- *)
PROGRAM PRG_Comms
// Comms task: lower priority than PRG_Control (e.g. 100 ms). One MQTT client for subscribing and
// publishing. Never touches Tags directly: commands go in through GVL_Tags.Commands, data comes out
// through GVL_Tags.PublishSnapshot, acknowledgements through GVL_Tags.Acks.
VAR CONSTANT
	TAGS_PER_CALL : INT := 250;         // spread a large build over several calls
	FULL_REFRESH_EVERY : UDINT := 60;   // every 60th message carries every tag
END_VAR
VAR
	BrokerUrl : STRING(64) := '192.168.50.240:1883';
	TopicData : STRING(64) := 'raw_data';
	TopicCommands : STRING(64) := 'plc_commands/CONC-BCNF-PLC';
	TopicAcks : STRING(64) := 'plc_acks/CONC-BCNF-PLC';

	MqttLink : MQTT.MQTT_IN_OUT;
	Subscriber : MQTT.MQTTSubscribe;
	Receiver : FB_CommandReceiver;
	Publisher : MQTT.MQTTPublish;
	AckPublisher : MQTT.MQTTPublish;
	IsInitialized : BOOL;
	ClientCallsMax : INT := 16;         // most client calls per scan while a message is in flight
	ClientBudgetUs : ULINT := 5000;     // ... and no more calls once this much time went into the client
	ClientCall : INT;
	ClientStartUs : ULINT;
	IsSendInFlight : BOOL;
	ConnectedEdge : R_TRIG;

	// Data publishing (PublishData, AppendTag, CommitSent, ForgetMessage)
	PublishTimer : TON;
	IsWaitingForSnapshot : BOOL;
	IsBuilding : BOOL;
	IsMessageReady : BOOL;              // built, waiting for the publisher to be armed
	IsRequested : BOOL;                 // send input of Publisher
	IsPublisherArmed : BOOL := TRUE;    // Publisher has seen send = FALSE since its last message
	IsBuildOk : BOOL;
	IsFullRefresh : BOOL;
	IsForceFullRefresh : BOOL := TRUE;  // the first message, and the next one after a reconnect or overflow
	SlowPublishEdge : R_TRIG;
	SlowPublishCount : UDINT;           // messages that took longer than the library's send time-out
	PublishCount : UDINT;
	NextTag : INT;
	LastTag : INT;
	Index : INT;
	Payload : STRING(32000);            // the generator sizes this from the table's worst-case message
	Used : UDINT;
	TagValue : REAL;
	ValueText : STRING(40);
	// Report-by-exception history: what the bridge last received, committed only after a message went out.
	LastSentValue : ARRAY[1..GVL_Tags.TAG_COUNT] OF REAL;
	LastSentQuality : ARRAY[1..GVL_Tags.TAG_COUNT] OF E_Quality;
	IsInMessage : ARRAY[1..GVL_Tags.TAG_COUNT] OF BOOL;

	// Acknowledgements (PublishAcks)
	Ack : ST_Command;
	AckLine : STRING(40);
	AckPayload : STRING(1000);
	AckUsed : UDINT;
	IsAckBatchReady : BOOL;             // a batch is built and not yet confirmed by the broker
	IsAckRequested : BOOL;
	IsAckPublisherArmed : BOOL := TRUE;
END_VAR
// ---- implementation ----
MqttLink.ClientID := 'CONC-BCNF-PLC';
// The client moves one 4 KB send buffer per two calls. While a message is in flight, call it again until
// ClientCallsMax calls or ClientBudgetUs; otherwise once, for keep-alive and receiving. This task's priority
// is below PRG_Control's, so the extra calls only use time control doesn't need.
IsSendInFlight := Publisher.sendActive OR AckPublisher.sendActive;
ClientStartUs := F_NowUs();
ClientCall := 0;
REPEAT
	MqttLink.clientFB(MQTT_IN_OUT := MqttLink, ENABLE := TRUE, URL := BrokerUrl, TIMEOUT := T#10S, TLS := FALSE);
	ClientCall := ClientCall + 1;
UNTIL ClientCall >= ClientCallsMax OR_ELSE NOT IsSendInFlight OR_ELSE F_NowUs() - ClientStartUs >= ClientBudgetUs
END_REPEAT
IF NOT IsInitialized THEN
	IsInitialized := TRUE;
	Subscriber.SetMqttInOut(MQTT_IN_OUT := MqttLink);
	Publisher.SetMqttInOut(MQTT_IN_OUT := MqttLink);
	AckPublisher.SetMqttInOut(MQTT_IN_OUT := MqttLink);
END_IF

Subscriber(Subscribe := TRUE, Topic := ADR(TopicCommands), QoSSubscribe := MQTT.QoS.AtLeastOnce,
	ExpectingString := TRUE, Callback := Receiver);
PublishData();
PublishAcks();

(* ---- PRG_Control.ApplyCommands.st ---- *)
// Action ApplyCommands (step 2): writable tags (setpoints, requests) are written here and nowhere else.
// Takes queued commands, checks them (CheckCommand), applies the accepted ones and answers every one.
// ---- implementation ----
// First scan: writable tags start from their configured defaults. Persisted setpoints, once added
// (a PERSISTENT copy owned by this step), are restored here instead.
IF NOT IsStarted THEN
	IsStarted := TRUE;
	FOR Index := 1 TO GVL_Tags.TAG_COUNT DO
		IF GVL_Tags.TagConfig[Index].IsWritable THEN
			GVL_Tags.Tags[Index].Value := GVL_Tags.TagConfig[Index].DefaultValue;
			GVL_Tags.Tags[Index].Quality := E_Quality.GOOD;
			GVL_Tags.Tags[Index].UpdatedAtMs := NowAtMs;
		END_IF
	END_FOR
END_IF

FOR Index := 1 TO MAX_COMMANDS_PER_SCAN DO
	IF NOT GVL_Tags.Commands.Pop(Item := Command) THEN
		EXIT;
	END_IF
	IsRetry := FALSE;
	IF Command.Result = E_CommandResult.PENDING THEN
		CheckCommand();
		IF NOT IsRetry THEN
			// The ledger holds every checked command with its answer, oldest replaced first. The generator sizes
			// it for all the commands the bridge may send within MAX_COMMAND_AGE_MS; a retry older than that
			// is TOO_OLD anyway. LedgerTooSmall counts entries replaced while still inside that window.
			IF Ledger[NextLedgerSlot].Id <> 0
					AND Ledger[NextLedgerSlot].SentAtMs + MAX_COMMAND_AGE_MS >= WallClockAtMs THEN
				LedgerTooSmall := LedgerTooSmall + 1;
			END_IF
			Ledger[NextLedgerSlot] := Command;
			NextLedgerSlot := (NextLedgerSlot + 1) MOD LEDGER_SIZE;
		END_IF
	END_IF
	IF IsRetry THEN
		RetriesAnswered := RetriesAnswered + 1;
	ELSIF Command.Result = E_CommandResult.ACCEPTED THEN
		GVL_Tags.Tags[Command.TagIndex].Value := Command.Value;
		GVL_Tags.Tags[Command.TagIndex].Quality := E_Quality.GOOD;
		GVL_Tags.Tags[Command.TagIndex].UpdatedAtMs := NowAtMs;
		GVL_Tags.Tags[Command.TagIndex].LastCommandSentAtMs := Command.SentAtMs;
		CommandsAccepted := CommandsAccepted + 1;
	ELSE
		CommandsRejected := CommandsRejected + 1;
	END_IF
	// A full Acks queue never holds a command back: a stop is applied even when its answer can't be queued.
	// The sender then times out and retries the same line, and the ledger answers it.
	IF NOT GVL_Tags.Acks.Push(Item := Command) THEN
		AcksDropped := AcksDropped + 1;
	END_IF
END_FOR

// A trip clears the start request, after the commands so a queued start can't undo it, and moves the trip
// time on for as long as the permit is missing. Uses last scan's permit; the output is already off through it.
IF NOT P_1502_Permit THEN
	GVL_Tags.Tags[GVL_Tags.TAG_P_1502_REQUEST].Value := 0.0;
	P_1502_TrippedAtMs := WallClockAtMs;
END_IF

(* ---- PRG_Control.CheckCommand.st ---- *)
// Action CheckCommand (part of step 2): sets Command.Result for a PENDING command. ACCEPTED means it may be
// applied. Range checks are written as NOT (inside) so that NaN and infinity count as outside.
// ---- implementation ----
// A retry is the identical line sent again: same id, tag, value and timestamp. It gets the first answer and
// is never applied twice. The same id with other content is a different command and is checked as new.
FOR Slot := 0 TO LEDGER_SIZE - 1 DO
	IF Ledger[Slot].Id = Command.Id AND Ledger[Slot].SentAtMs = Command.SentAtMs
			AND Ledger[Slot].TagIndex = Command.TagIndex AND Ledger[Slot].Value = Command.Value THEN
		Command.Result := Ledger[Slot].Result;
		IsRetry := TRUE;
		RETURN;
	END_IF
END_FOR

IF Command.TagIndex = 0 THEN
	Command.Result := E_CommandResult.UNKNOWN_TAG;
ELSIF NOT GVL_Tags.TagConfig[Command.TagIndex].IsWritable THEN
	Command.Result := E_CommandResult.NOT_WRITABLE;
ELSIF NOT (Command.Value >= GVL_Tags.TagConfig[Command.TagIndex].MinValue
		AND Command.Value <= GVL_Tags.TagConfig[Command.TagIndex].MaxValue) THEN
	Command.Result := E_CommandResult.OUT_OF_RANGE;
ELSIF GVL_Tags.TagConfig[Command.TagIndex].Kind = E_TagKind.BOOL_TAG
		AND Command.Value <> 0.0 AND Command.Value <> 1.0 THEN
	Command.Result := E_CommandResult.OUT_OF_RANGE;
// Converted only once the value is inside the tag's range, which the generator keeps inside DINT.
ELSIF GVL_Tags.TagConfig[Command.TagIndex].Kind = E_TagKind.INT_TAG
		AND_THEN Command.Value <> DINT_TO_REAL(REAL_TO_DINT(Command.Value)) THEN
	Command.Result := E_CommandResult.OUT_OF_RANGE;
ELSIF WallClockAtMs < MIN_PLAUSIBLE_WALL_CLOCK_MS THEN
	Command.Result := E_CommandResult.CLOCK_NOT_SYNCED;
ELSIF Command.SentAtMs > WallClockAtMs + MAX_FUTURE_SKEW_MS
		OR Command.SentAtMs + MAX_COMMAND_AGE_MS < WallClockAtMs
		OR (Command.ReceivedAtMs < NowAtMs AND NowAtMs - Command.ReceivedAtMs > MAX_QUEUE_AGE_MS) THEN
	Command.Result := E_CommandResult.TOO_OLD;
// Every timestamp comes from one clock, the bridge's (the only command sender), so they can be ordered.
ELSIF Command.SentAtMs < GVL_Tags.Tags[Command.TagIndex].LastCommandSentAtMs THEN
	Command.Result := E_CommandResult.OUT_OF_ORDER;      // a newer command for this tag already applied
// A start must be sent after the permit came back, with the clock skew as margin. A start that was queued
// or delayed across a trip, or retried after one, is refused.
ELSIF Command.TagIndex = GVL_Tags.TAG_P_1502_REQUEST AND Command.Value > 0.5
		AND (NOT P_1502_Permit OR Command.SentAtMs <= P_1502_TrippedAtMs + MAX_FUTURE_SKEW_MS) THEN
	Command.Result := E_CommandResult.INTERLOCKED;
ELSE
	Command.Result := E_CommandResult.ACCEPTED;
END_IF

(* ---- PRG_Control.CollectBusInputs.st ---- *)
// Action CollectBusInputs (start of step 1): device values and health from the bus task. A source the bus task
// was updating when this scan started (SourceWriting) keeps last scan's values; it is complete next scan.
// ---- implementation ----
FOR Index := 1 TO GVL_Tags.SOURCE_COUNT DO
	IF GVL_Bus.IsBusSource[Index] AND NOT GVL_Bus.SourceWriting[Index] THEN
		GVL_Tags.SourceIsHealthy[Index] := GVL_Bus.SourceHealthy[Index];
		GVL_Tags.SourceUpdatedAtMs[Index] := GVL_Bus.SourceLastGoodMs[Index];
	END_IF
END_FOR
FOR Index := 1 TO GVL_Tags.TAG_COUNT DO
	Slot := GVL_Tags.TagConfig[Index].Source;
	IF GVL_Bus.IsBusSource[Slot] AND NOT GVL_Bus.SourceWriting[Slot] THEN
		GVL_Tags.RawInputs[Index] := GVL_Bus.Raw[Index];
	END_IF
END_FOR

(* ---- PRG_Control.ComputeValues.st ---- *)
// Action ComputeValues (step 3): engineering value and final quality for every input tag: the source's
// quality, downgraded to INVALID when the value is out of range or not a number. Derived values (recovery %,
// rejection %) go here too, computed only when their inputs are GOOD and the divisor is not zero.
// ---- implementation ----
FOR Index := 1 TO GVL_Tags.TAG_COUNT DO
	IF NOT GVL_Tags.TagConfig[Index].IsWritable THEN
		GVL_Tags.Tags[Index].Value := GVL_Tags.Tags[Index].Raw * GVL_Tags.TagConfig[Index].Scale
			+ GVL_Tags.TagConfig[Index].Offset;
		GVL_Tags.Tags[Index].Quality := GVL_Tags.Tags[Index].SourceQuality;
		// Written as NOT (inside the range) so that NaN and infinity, which fail every comparison, are INVALID.
		IF GVL_Tags.Tags[Index].Quality = E_Quality.GOOD
				AND NOT (GVL_Tags.Tags[Index].Value >= GVL_Tags.TagConfig[Index].MinValue
					AND GVL_Tags.Tags[Index].Value <= GVL_Tags.TagConfig[Index].MaxValue) THEN
			GVL_Tags.Tags[Index].Quality := E_Quality.INVALID;
		END_IF
	END_IF
END_FOR

(* ---- PRG_Control.EvaluateAlarms.st ---- *)
// Action EvaluateAlarms (step 4). One alarm shown; in the full design alarms are rows in a generated
// table (tag, setpoint tag, direction, hysteresis, delay, priority) evaluated in a loop.
// ---- implementation ----
// HH alarm with hysteresis. A value or a setpoint that can't be trusted counts as an alarm (fail safe).
IF GVL_Tags.Tags[GVL_Tags.TAG_AIT_1508].Quality <> E_Quality.GOOD
		OR GVL_Tags.Tags[GVL_Tags.TAG_AIT_1508_HH_SP].Quality <> E_Quality.GOOD THEN
	AIT_1508_HH := TRUE;
ELSIF GVL_Tags.Tags[GVL_Tags.TAG_AIT_1508].Value >= GVL_Tags.Tags[GVL_Tags.TAG_AIT_1508_HH_SP].Value THEN
	AIT_1508_HH := TRUE;
ELSIF GVL_Tags.Tags[GVL_Tags.TAG_AIT_1508].Value
		< GVL_Tags.Tags[GVL_Tags.TAG_AIT_1508_HH_SP].Value - ALARM_HYSTERESIS THEN
	AIT_1508_HH := FALSE;
END_IF

// A remote E-stop is active unless it is positively reported clear: an untrusted signal, or one that has
// stopped arriving, counts as a stop. NOT (< 0.5) also treats NaN as a stop.
LSS_E_STOP_ACTIVE := NOT (GVL_Tags.Tags[GVL_Tags.TAG_LSS_E_STOP].Value < 0.5)
	OR GVL_Tags.Tags[GVL_Tags.TAG_LSS_E_STOP].Quality <> E_Quality.GOOD;

(* ---- PRG_Control.ReadInputs.st ---- *)
// Action ReadInputs (step 1): raw values and the quality of their source. A failed or silent source keeps
// its last good raw value, marked, instead of whatever the I/O image holds. Requests and setpoints are not
// inputs: they only change through ApplyCommands.
// ---- implementation ----
CollectBusInputs();     // devices on the Modbus lines (bus task)
FOR Index := 1 TO GVL_Tags.TAG_COUNT DO
	IF NOT GVL_Tags.TagConfig[Index].IsWritable THEN
		IF NOT GVL_Tags.SourceIsHealthy[GVL_Tags.TagConfig[Index].Source] THEN
			GVL_Tags.Tags[Index].SourceQuality := E_Quality.COMM_FAIL;       // local I/O diagnostics too
		ELSIF GVL_Tags.TagConfig[Index].Source = 0 THEN
			GVL_Tags.Tags[Index].Raw := GVL_Tags.RawInputs[Index];
			GVL_Tags.Tags[Index].SourceQuality := E_Quality.GOOD;
			GVL_Tags.Tags[Index].UpdatedAtMs := NowAtMs;
		ELSIF GVL_Tags.SourceUpdatedAtMs[GVL_Tags.TagConfig[Index].Source] = 0 THEN
			GVL_Tags.Tags[Index].SourceQuality := E_Quality.INIT;            // no sample since start-up
		ELSIF GVL_Tags.SourceUpdatedAtMs[GVL_Tags.TagConfig[Index].Source] < NowAtMs
				AND NowAtMs - GVL_Tags.SourceUpdatedAtMs[GVL_Tags.TagConfig[Index].Source]
					> TIME_TO_ULINT(GVL_Tags.TagConfig[Index].StaleAfter) THEN
			GVL_Tags.Tags[Index].SourceQuality := E_Quality.STALE;
		ELSE
			GVL_Tags.Tags[Index].Raw := GVL_Tags.RawInputs[Index];
			GVL_Tags.Tags[Index].SourceQuality := E_Quality.GOOD;
			GVL_Tags.Tags[Index].UpdatedAtMs := GVL_Tags.SourceUpdatedAtMs[GVL_Tags.TagConfig[Index].Source];
		END_IF
	END_IF
END_FOR

(* ---- PRG_Control.ServeSnapshot.st ---- *)
// Action ServeSnapshot (step 7): when the comms task asks (SnapshotRequest moved on), copy the whole tag
// table at once, inside this task, so a published message never mixes values from different scans.
// ---- implementation ----
IF GVL_Tags.SnapshotSequence <> GVL_Tags.SnapshotRequest THEN
	GVL_Tags.PublishSnapshot := GVL_Tags.Tags;
	GVL_Tags.SnapshotSequence := GVL_Tags.SnapshotRequest;
END_IF

(* ---- PRG_Control.st ---- *)
PROGRAM PRG_Control
// Control task: high priority, fixed interval (e.g. 50 ms). Runs the same pipeline every scan. Each step
// writes only its own results and reads only what the steps before it produced, so the order is the design.
VAR CONSTANT
	MAX_COMMANDS_PER_SCAN : INT := 10;  // bound the command work per scan; the rest waits in the queue
	MAX_COMMAND_AGE_MS : ULINT := 10000;
	MAX_FUTURE_SKEW_MS : ULINT := 2000; // a command dated further ahead than this is rejected
	MAX_QUEUE_AGE_MS : ULINT := 2000;   // ... and so is one that waited longer than this in the queue
	MIN_PLAUSIBLE_WALL_CLOCK_MS : ULINT := 1700000000000;  // before 2023-11: the RTC is not synchronized
	LEDGER_SIZE : INT := 64;            // answered commands remembered for retries; see ApplyCommands
	ALARM_HYSTERESIS : REAL := 0.1;
END_VAR
VAR
	NowAtMs : ULINT;                    // monotonic, for ages
	WallClockAtMs : ULINT;              // real-time clock, for command timestamps
	IsStarted : BOOL;
	Index : INT;
	Slot : INT;
	Command : ST_Command;

	// Command bookkeeping (ApplyCommands, CheckCommand)
	Ledger : ARRAY[0..LEDGER_SIZE - 1] OF ST_Command;
	NextLedgerSlot : INT;
	IsRetry : BOOL;

	// Alarms (EvaluateAlarms)
	AIT_1508_HH : BOOL;
	LSS_E_STOP_ACTIVE : BOOL;

	// Permissives (EvaluatePermissives)
	P_1502_Permit : BOOL;
	IsBypassActive : BOOL;
	P_1502_TrippedAtMs : ULINT;         // wall clock, last scan without the permit (ApplyCommands)
	BypassUntilMs : ULINT;              // a remote bypass expires; 0 = none (command path not in the skeleton)
	LocalBypassEnable : BOOL;           // key switch input: a remote bypass only works with it on

	// Diagnostics
	CommandsAccepted : UDINT;
	CommandsRejected : UDINT;
	RetriesAnswered : UDINT;
	AcksDropped : UDINT;
	LedgerTooSmall : UDINT;
END_VAR
// ---- implementation ----
NowAtMs := F_NowMs();
WallClockAtMs := F_WallClockMs();

ReadInputs();          // 1. I/O and bus values -> Tags[].Raw; quality from source health and age
ApplyCommands();       // 2. queued remote commands -> validated setpoints and requests, acknowledged
ComputeValues();       // 3. scaling, range checks, derived values
EvaluateAlarms();      // 4. alarm bits from values, quality and setpoints
EvaluatePermissives(); // 5. interlocks: what is allowed to run
WriteOutputs();        // 6. output := request AND permit; the only place outputs are written
ServeSnapshot();       // 7. a consistent copy of Tags for the comms task, when it asks
